// TIA Portal project "2026_10_06_Lavorazione_Olive" (V15)

(* hardware
DEVICE "S7-1200 station_1"  S7-1200 Station
   slot 0: "Telaio di montaggio_0"  S7-1200 Rack  Rack  V1.0
   slot 1: "PLC_1"  CPU 1215C DC/DC/DC  6ES7 215-1AG40-0XB0  V4.2
*)

// ===== PLC "PLC_1"  CPU 1215C DC/DC/DC =====

VAR_GLOBAL   // PLC tag table "Tabella delle variabili standard"
   "SP" AT %I0.0 : Bool;   // Sensore di presenza olive
   "ST" AT %IW64 : Word;   // Sensore analogico di temperatura
   "KM1" AT %Q0.0 : Bool;   // Motore M1 del frangitore
   "KM2" AT %Q0.1 : Bool;   // Motore M2 del granulatore
   "KM3" AT %Q0.2 : Bool;   // Motore M3 dell'elettropompa
   "KER" AT %Q0.3 : Bool;   // Elementi riscaldanti
   "HLP" AT %Q0.4 : Bool;   // Lampada di segnalazione presenza
   "HLL" AT %Q0.5 : Bool;   // Lampada lampeggio sistema acceso
   "T_Norm" AT %MD3 : Real;   // Temperatura normalizzata
   "T_Real" AT %MD4 : Real;   // Temperatura reale
   "P0" AT %M20.0 : Bool;   // Attesa presenza prodotto
   "P1" AT %M20.1 : Bool;   // Avvio M1, M2, M3
   "P2" AT %M20.2 : Bool;   // Attesa T_F (5 minuti)
   "P3" AT %M20.3 : Bool;   // Attesa T_G (40 minuti)
   "P_T" AT %M20.4 : Bool;   // Stato attivazione elementi riscaldanti
   "Clock_Byte" AT %MB0 : Byte;
   "Clock_10Hz" AT %M0.0 : Bool;
   "Clock_5Hz" AT %M0.1 : Bool;
   "Clock_2.5Hz" AT %M0.2 : Bool;
   "Clock_2Hz" AT %M0.3 : Bool;
   "Clock_1.25Hz" AT %M0.4 : Bool;
   "Clock_1Hz" AT %M0.5 : Bool;
   "Clock_0.625Hz" AT %M0.6 : Bool;
   "Clock_0.5Hz" AT %M0.7 : Bool;
   "System_Byte" AT %MB1 : Byte;
   "FirstScan" AT %M1.0 : Bool;
   "DiagStatusUpdate" AT %M1.1 : Bool;
   "AlwaysTRUE" AT %M1.2 : Bool;
   "AlwaysFALSE" AT %M1.3 : Bool;
   "P" AT %MW30 : Int;   // Variabile di stato
END_VAR

// folder: System blocks/Program resources

DATA_BLOCK "T_F"   // DB1
{ S7_Optimized_Access := 'TRUE' }
AUTHOR : Simatic
FAMILY : IEC
NAME : IEC_TMR
VERSION : 1.0
// stored: InstanceOfName IEC_TIMER
"IEC_TIMER"
BEGIN
END_DATA_BLOCK

DATA_BLOCK "T_G"   // DB2
{ S7_Optimized_Access := 'TRUE' }
AUTHOR : Simatic
FAMILY : IEC
NAME : IEC_TMR
VERSION : 1.0
// stored: InstanceOfName IEC_TIMER
"IEC_TIMER"
BEGIN
END_DATA_BLOCK

// folder: (top level)

FUNCTION "Controllo" : Void   // FC1, LAD
{ S7_Optimized_Access := 'TRUE' }
VERSION : 0.1
BEGIN

REGION Network 1: Avvio sistema
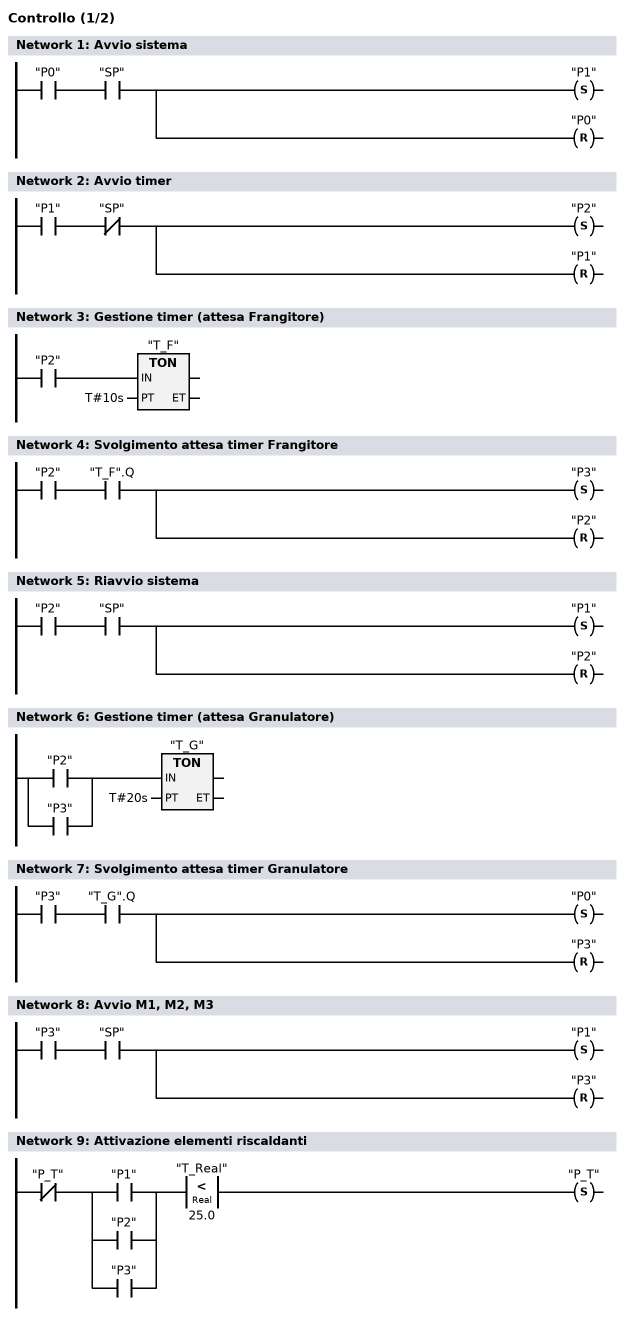
   RUNG wire#powerrail
      Contact( "P0" )
      Contact( "SP" )
      wire#w1
      S_Coil( "P1" )
   END_RUNG
   RUNG wire#w1
      R_Coil( "P0" )
   END_RUNG
   // the same network as SCL:
   IF "P0" AND "SP" THEN
       "P1" := TRUE;
       "P0" := FALSE;
   END_IF;
END_REGION

REGION Network 2: Avvio timer
   RUNG wire#powerrail
      Contact( "P1" )
      I_Contact( "SP" )
      wire#w1
      S_Coil( "P2" )
   END_RUNG
   RUNG wire#w1
      R_Coil( "P1" )
   END_RUNG
   // the same network as SCL:
   IF "P1" AND NOT "SP" THEN
       "P2" := TRUE;
       "P1" := FALSE;
   END_IF;
END_REGION

REGION Network 3: Gestione timer (attesa Frangitore)
   "T_F".TON(IN := "P2", PT := T#10s);
END_REGION

REGION Network 4: Svolgimento attesa timer Frangitore
   RUNG wire#powerrail
      Contact( "P2" )
      Contact( "T_F".Q )
      wire#w1
      S_Coil( "P3" )
   END_RUNG
   RUNG wire#w1
      R_Coil( "P2" )
   END_RUNG
   // the same network as SCL:
   IF "P2" AND "T_F".Q THEN
       "P3" := TRUE;
       "P2" := FALSE;
   END_IF;
END_REGION

REGION Network 5: Riavvio sistema
   RUNG wire#powerrail
      Contact( "P2" )
      Contact( "SP" )
      wire#w1
      S_Coil( "P1" )
   END_RUNG
   RUNG wire#w1
      R_Coil( "P2" )
   END_RUNG
   // the same network as SCL:
   IF "P2" AND "SP" THEN
       "P1" := TRUE;
       "P2" := FALSE;
   END_IF;
END_REGION

REGION Network 6: Gestione timer (attesa Granulatore)
   "T_G".TON(IN := "P2" OR "P3", PT := T#20s);
END_REGION

REGION Network 7: Svolgimento attesa timer Granulatore
   RUNG wire#powerrail
      Contact( "P3" )
      Contact( "T_G".Q )
      wire#w1
      S_Coil( "P0" )
   END_RUNG
   RUNG wire#w1
      R_Coil( "P3" )
   END_RUNG
   // the same network as SCL:
   IF "P3" AND "T_G".Q THEN
       "P0" := TRUE;
       "P3" := FALSE;
   END_IF;
END_REGION

REGION Network 8: Avvio M1, M2, M3
   RUNG wire#powerrail
      Contact( "P3" )
      Contact( "SP" )
      wire#w1
      S_Coil( "P1" )
   END_RUNG
   RUNG wire#w1
      R_Coil( "P3" )
   END_RUNG
   // the same network as SCL:
   IF "P3" AND "SP" THEN
       "P1" := TRUE;
       "P3" := FALSE;
   END_IF;
END_REGION

REGION Network 9: Attivazione elementi riscaldanti
   RUNG wire#powerrail
      I_Contact( "P_T" )
      wire#w1
      Contact( "P1" )
      wire#w2
      { S7_Templates := "SrcType := Real" } LT_Contact(in1 := "T_Real", in2 := 25.0)
      S_Coil( "P_T" )
   END_RUNG
   RUNG wire#w1
      Contact( "P2" )
   END_RUNG wire#w2
   RUNG wire#w1
      Contact( "P3" )
   END_RUNG wire#w2
   // the same network as SCL:
   IF NOT "P_T" AND ("P1" OR "P2" OR "P3") AND ("T_Real" < 25.0) THEN "P_T" := TRUE; END_IF;
END_REGION

REGION Network 10: Disattivazione elementi riscaldanti
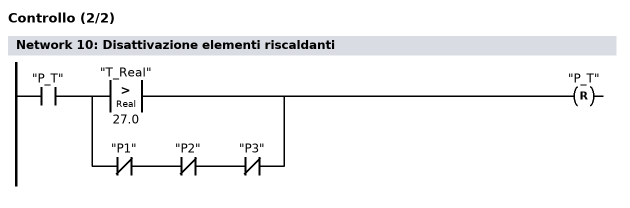
   RUNG wire#powerrail
      Contact( "P_T" )
      wire#w1
      { S7_Templates := "SrcType := Real" } GT_Contact(in1 := "T_Real", in2 := 27.0)
      wire#w2
      R_Coil( "P_T" )
   END_RUNG
   RUNG wire#w1
      I_Contact( "P1" )
      I_Contact( "P2" )
      I_Contact( "P3" )
   END_RUNG wire#w2
   // the same network as SCL:
   IF "P_T" AND (("T_Real" > 27.0) OR (NOT "P1" AND NOT "P2" AND NOT "P3")) THEN "P_T" := FALSE; END_IF;
END_REGION
END_FUNCTION

FUNCTION "Comando" : Void   // FC2, LAD
{ S7_Optimized_Access := 'TRUE' }
VERSION : 0.1
BEGIN

REGION Network 1: Motore M1 del frangitore
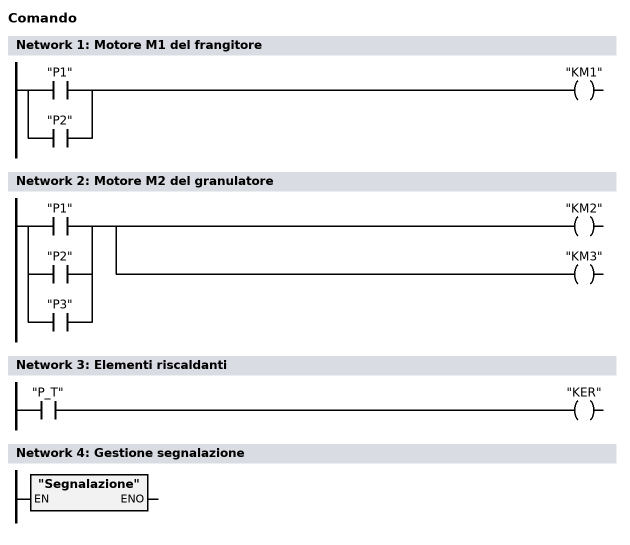
   RUNG wire#powerrail
      Contact( "P1" )
      wire#w1
      Coil( "KM1" )
   END_RUNG
   RUNG wire#powerrail
      Contact( "P2" )
   END_RUNG wire#w1
   // the same network as SCL:
   "KM1" := "P1" OR "P2";
END_REGION

REGION Network 2: Motore M2 del granulatore
   RUNG wire#powerrail
      Contact( "P1" )
      wire#w1
      Coil( "KM2" )
   END_RUNG
   RUNG wire#powerrail
      Contact( "P2" )
   END_RUNG wire#w1
   RUNG wire#powerrail
      Contact( "P3" )
   END_RUNG wire#w1
   RUNG wire#w1
      Coil( "KM3" )
   END_RUNG
   // the same network as SCL:
   "KM2" := "P1" OR "P2" OR "P3";
   "KM3" := "KM2";
END_REGION

REGION Network 3: Elementi riscaldanti
   RUNG wire#powerrail
      Contact( "P_T" )
      Coil( "KER" )
   END_RUNG
   // the same network as SCL:
   "KER" := "P_T";
END_REGION

REGION Network 4: Gestione segnalazione
   RUNG wire#powerrail
      "Segnalazione"()
   END_RUNG
   // the same network as SCL:
   "Segnalazione"();
END_REGION
END_FUNCTION

FUNCTION "Segnalazione" : Void   // FC3, LAD
{ S7_Optimized_Access := 'TRUE' }
VERSION : 0.1
BEGIN

REGION Network 1: Lampada di segnalazione presenza
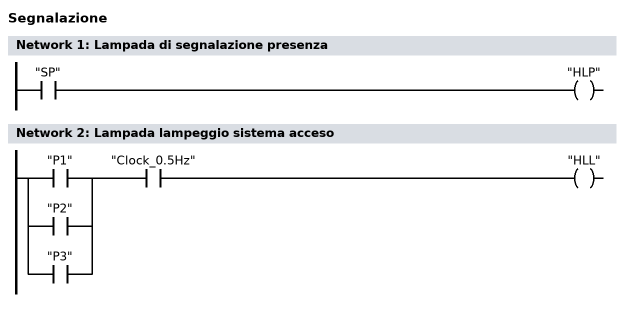
   RUNG wire#powerrail
      Contact( "SP" )
      Coil( "HLP" )
   END_RUNG
   // the same network as SCL:
   "HLP" := "SP";
END_REGION

REGION Network 2: Lampada lampeggio sistema acceso
   RUNG wire#powerrail
      Contact( "P1" )
      wire#w1
      Contact( "Clock_0.5Hz" )
      Coil( "HLL" )
   END_RUNG
   RUNG wire#powerrail
      Contact( "P2" )
   END_RUNG wire#w1
   RUNG wire#powerrail
      Contact( "P3" )
   END_RUNG wire#w1
   // the same network as SCL:
   "HLL" := ("P1" OR "P2" OR "P3") AND "Clock_0.5Hz";
END_REGION
END_FUNCTION

FUNCTION "Temperatura" : Void   // FC4, LAD
{ S7_Optimized_Access := 'TRUE' }
VERSION : 0.1
BEGIN

REGION Network 1: Trascrizione con blocco NORM
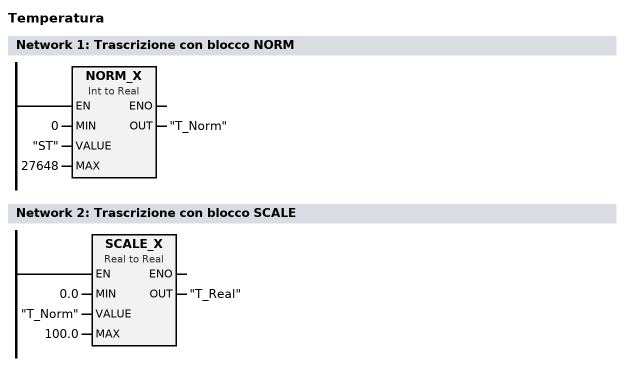
   RUNG wire#powerrail
      { S7_Templates := "[SrcType := Int, DestType := Real]" } Normalize(min := 0, value := "ST", max := 27648, out => "T_Norm")
   END_RUNG
   // the same network as SCL:
   "T_Norm" := NORM_X(MIN := 0, VALUE := "ST", MAX := 27648);
END_REGION

REGION Network 2: Trascrizione con blocco SCALE
   RUNG wire#powerrail
      { S7_Templates := "[SrcType := Real, DestType := Real]" } Scale(min := 0.0, value := "T_Norm", max := 100.0, out => "T_Real")
   END_RUNG
   // the same network as SCL:
   "T_Real" := SCALE_X(MIN := 0.0, VALUE := "T_Norm", MAX := 100.0);
END_REGION
END_FUNCTION

ORGANIZATION_BLOCK "Main"   // OB1, LAD, ProgramCycle
TITLE = "Main Program Sweep (Cycle)"
{ S7_Optimized_Access := 'TRUE' }
VERSION : 0.1
   VAR_INPUT
      Initial_Call : Bool;   // Initial call of this OB
      Remanence : Bool;   // =True, if remanent data are available
   END_VAR
BEGIN

REGION Network 1: FC misurazione temperatura
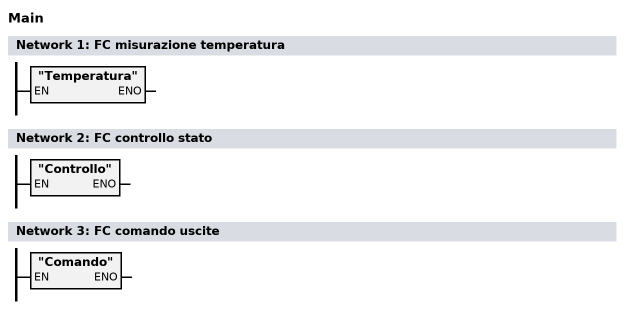
   RUNG wire#powerrail
      "Temperatura"()
   END_RUNG
   // the same network as SCL:
   "Temperatura"();
END_REGION

REGION Network 2: FC controllo stato
   RUNG wire#powerrail
      "Controllo"()
   END_RUNG
   // the same network as SCL:
   "Controllo"();
END_REGION

REGION Network 3: FC comando uscite
   RUNG wire#powerrail
      "Comando"()
   END_RUNG
   // the same network as SCL:
   "Comando"();
END_REGION
END_ORGANIZATION_BLOCK

ORGANIZATION_BLOCK "Startup"   // OB100, LAD, Startup
TITLE = "Complete Restart"
{ S7_Optimized_Access := 'TRUE' }
VERSION : 0.1
   VAR_INPUT
      LostRetentive : Bool;   // True if retentive data are lost
      LostRTC : Bool;   // True if date and time are lost
   END_VAR
BEGIN

REGION Network 1: Reset stato iniziale
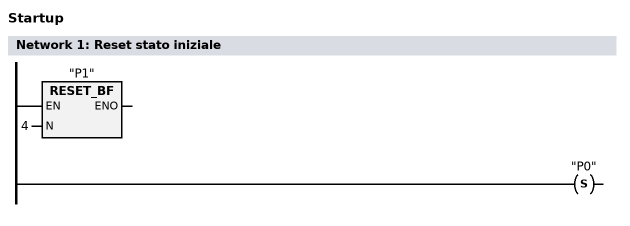
   // no SCL statement known for RBitfield: written as a call
   RESET_BF(operand := "P1", n := 4);
   "P0" := TRUE;
END_REGION
END_ORGANIZATION_BLOCK